Staubli VAL3: actItem.pjx

--- actItem.pjx ---
Parameters version=s8.10.3Cs9_BS2093 stackSize=5000 millimeterUnit=true
Data file=actItem.dtx
Type name=actionItem path=Disk://source/template/actionItem/actionItem.pjx

--- actItem.dtx ---
public string sComment
public actionItem aActItem[6]
  [0]
    num nIOindex
    num nboolValue
    num nPulseValue
    string sIOtype
    string sValue
    bool bActive
  [1]
    num nIOindex
    num nboolValue
    num nPulseValue
    string sIOtype
    string sValue
    bool bActive
  [2]
    num nIOindex
    num nboolValue
    num nPulseValue
    string sIOtype
    string sValue
    bool bActive
  [3]
    num nIOindex
    num nboolValue
    num nPulseValue
    string sIOtype
    string sValue
    bool bActive
  [4]
    num nIOindex
    num nboolValue
    num nPulseValue
    string sIOtype
    string sValue
    bool bActive
  [5]
    num nIOindex
    num nboolValue
    num nPulseValue
    string sIOtype
    string sValue
    bool bActive
